RoboDK station: Celda_Soldadura_Estator_Grupo4_v03.rdk

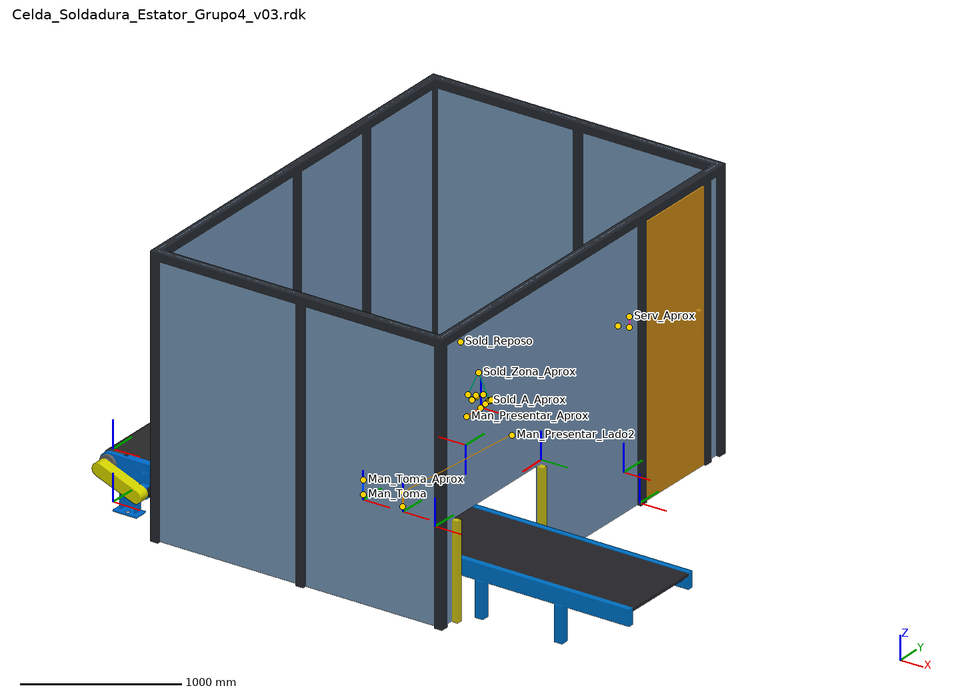
[picture v0: the station drawn from its stored meshes, robots at their saved joint values, targets as dots, program paths as lines]
Station Celda_Soldadura_Estator_Grupo4_v03 (saved by RoboDK 6.1.1). Poses are relative to the parent item; angles as X-Y-Z fixed-axis rotations.
Station parameters (name, value as stored): PIEZA_EN_TOMA, 0, PIEZA_PRESENTADA, 0, ARCO_TIG, 0, SOLDADURA_TERMINADA, 0
  - frame Frame_Celda at (0, 0, 0) mm
    - frame Base_Manipulador_IRB1200 at (0, 0, 0) mm
      - robot ABB IRB 1200-7/0.7: 6 axes, payload 7 kg, reach 703 mm, repeatability 0.02 mm, weight 54 kg
          modified DH rows (alpha deg, a mm, theta deg, d mm): 0, 0, 0, 399; -90, 0, -90, 0; 0, 350, 0, 0; -90, 42, 0, 351; 90, 0, 0, 0; -90, 0, 180, 82
          joint limits [-170, -100, -200, -270, -130, -360] to [170, 135, 70, 270, 130, 360]; home [0, 0, 0, 0, 0, 0]; saved at [0, -20, 30, 0, 80, 0]
        - frame RobotiQ 2F-85 Gripper (Mechanism) Base at (0, 0, 0) mm
          - robot Pinza_2F85 (model RobotiQ 2F85): 1 axes, payload 5 kg
              joint limits [0] to [85]; home [85]; saved at [0]
        - tool TCP_Pinza, TCP at (0, 0, 150) mm
    - frame Base_Soldador_CRB1300 at (0, 1150, 0) mm, rotated rx 0 ry 0 rz -90 deg
      - robot ABB CRB 1300-10/1.15: 6 axes
          modified DH rows (alpha deg, a mm, theta deg, d mm): 0, 0, 0, 544; -90, 150, -90, 0; 0, 575, 0, 0; -90, 40, 0, 425; 90, 0, 0, 0; -90, 0, 180, 90
          joint limits [-180, -95, -210, -230, -130, -242] to [180, 155, 65, 230, 130, 242]; home [0, 0, 0, 0, 0, 0]; saved at [0, -10, 10, 0, 60, 0]
        - tool Antorcha_TIG, TCP at (0, 0, 207) mm, size 80 x 80 x 207 mm, geometry from antorcha_tig.stl
    - frame Base_Cinta_Pasante at (-1830, -860, 0) mm
      - robot Cinta_Pasante: 1 axes
          modified DH rows (alpha deg, a mm, theta deg, d mm): 0, 0, 0, 0 linear
          base shift (0, 0, 0) mm, rotated rx 0 ry 90 rz 0 deg
          joint limits [-900000] to [900000]; home [0]; saved at [0]
        - frame Frame_Banda at (0, 0, 0) mm
          - frame Frame_Piezas_Soldadas at (0, 0, 0) mm
          - object Estator_1 at (1680, 300, 0) mm, size 105 x 105 x 55 mm, geometry from paquete_estator.stl
          - object Estator_2 at (1380, 300, 0) mm, size 105 x 105 x 55 mm, geometry from paquete_estator.stl
          - object Estator_3 at (1080, 300, 0) mm, size 105 x 105 x 55 mm, geometry from paquete_estator.stl
          - object Estator_4 at (780, 300, 0) mm, size 105 x 105 x 55 mm, geometry from paquete_estator.stl
    - object Sensor_Pieza_En_Toma at (-150, -900, 396.5) mm, rotated rx 0 ry 0 rz 90 deg, size 683.3 x 45.2 x 12.5 mm, geometry from Laser-Sensor.stl
    - object Estacion_Servicio_Antorcha at (520, 1300, 0) mm, size 250 x 250 x 1000 mm, geometry from estacion_servicio_antorcha.stl
    - frame Frame_Cerramiento at (0, 0, 0) mm
      - frame Bisagra_Puerta at (850, 1000, 0) mm
        - object Puerta at (0, 0, 0) mm, size 60 x 700 x 1920 mm, geometry from puerta.stl
      - object Cerramiento_Estructura at (0, 0, 0) mm, size 2210 x 3060 x 2000 mm, geometry from cerramiento_estructura_v03.stl
      - object Cerramiento_Paneles at (0, 0, 0) mm, size 2154 x 3004 x 2000 mm, geometry from cerramiento_paneles_v03.stl
      - object Cortina_Luz_Entrada at (-1330, 0, 0) mm, size 40 x 960 x 700 mm, geometry from cortina_luz_cinta.stl
      - object Cortina_Luz_Salida at (880, 0, 0) mm, size 40 x 960 x 700 mm, geometry from cortina_luz_cinta.stl
    - frame Frame_Soldadura at (0, 500, 620) mm
      - target Man_Presentar_Aprox (Cartesian target) at (0, -157.5, 0) mm, rotated rx -90 ry 0 rz 0 deg; joints [0, 0, 0, 0, 0, 0] of ABB IRB 1200-7/0.7
      - target Man_Presentar_Lado1 (Cartesian target) at (0, -7.5, 0) mm, rotated rx -90 ry 0 rz 0 deg; joints [0, 0, 0, 0, 0, 0] of ABB IRB 1200-7/0.7
      - target Man_Presentar_Lado2 (joint target) at (583, -500, 171) mm, rotated rx 0 ry 90 rz 0 deg; joints [90, -11.774, 38.724, 0, -26.95, 90] of ABB IRB 1200-7/0.7
      - target Man_Presentar_Aprox_Lado2 (joint target) at (583, -500, 171) mm, rotated rx 0 ry 90 rz 0 deg; joints [90, -43.636, 55.703, 0, -12.068, 90] of ABB IRB 1200-7/0.7
      - target Sold_Zona_Aprox (Cartesian target) at (0, -26.5, 250) mm, rotated rx 180 ry 0 rz 90 deg; joints [103.36, 41.617, 53.414, 0, -5.031, 103.36] of ABB CRB 1300-10/1.15
      - target Sold_A_Aprox (Cartesian target) at (78.2, -26.5, 78.2) mm, rotated rx -135 ry 0 rz 90 deg; joints [98.688, 74.302, 5.58, 7.491, 55.018, 91.856] of ABB CRB 1300-10/1.15
      - target Sold_A_Inicio (Cartesian target) at (49.91, -26.5, 49.91) mm, rotated rx -135 ry 0 rz 90 deg; joints [98.998, 76.411, 8.063, 8.245, 50.464, 91.119] of ABB CRB 1300-10/1.15
      - target Sold_A_Fin (Cartesian target) at (49.91, 26.5, 49.91) mm, rotated rx -135 ry 0 rz 90 deg; joints [102.751, 76.611, 6.557, 11.474, 51.681, 91.918] of ABB CRB 1300-10/1.15
      - target Sold_Transicion_Medio (Cartesian target) at (0, 26.5, 80) mm, rotated rx 180 ry 0 rz 90 deg; joints [108.748, 65.119, 46.933, 0, -22.052, 108.748] of ABB CRB 1300-10/1.15
      - target Sold_B_Inicio (Cartesian target) at (-49.91, 26.5, 49.91) mm, rotated rx 135 ry 0 rz 90 deg; joints [124.163, 102.688, 60.997, 205.222, 111.278, -54.665] of ABB CRB 1300-10/1.15
      - target Sold_B_Fin (Cartesian target) at (-49.91, -26.5, 49.91) mm, rotated rx 135 ry 0 rz 90 deg; joints [115.401, 107.202, 62.682, 200.569, 120.307, -60.716] of ABB CRB 1300-10/1.15
      - target Sold_B_Retiro (Cartesian target) at (-78.2, -26.5, 78.2) mm, rotated rx 135 ry 0 rz 90 deg; joints [-61.951, -75.264, -208.995, 23.114, 57.885, -82.141] of ABB CRB 1300-10/1.15
      - target Sold_A_Salida (Cartesian target) at (56.57, 26.5, 56.57) mm, rotated rx -135 ry 0 rz 90 deg; joints [102.647, 76.107, 6.003, 11.22, 52.72, 92.165] of ABB CRB 1300-10/1.15
      - target Sold_B_Entrada (Cartesian target) at (-56.57, 26.5, 56.57) mm, rotated rx 135 ry 0 rz 90 deg; joints [124.856, 103.181, 62.152, 205.935, 112.476, -53.248] of ABB CRB 1300-10/1.15
    - frame Frame_Toma_Cinta at (-150, -560, 366.5) mm
      - target Man_Toma_Aprox (Cartesian target) at (0, 0, 135) mm, rotated rx 180 ry 0 rz 0 deg; joints [0, 0, 0, 0, 0, 0] of ABB IRB 1200-7/0.7
      - target Man_Toma (Cartesian target) at (0, 0, 35) mm, rotated rx 180 ry 0 rz 0 deg; joints [0, 0, 0, 0, 0, 0] of ABB IRB 1200-7/0.7
    - frame Frame_Servicio at (520, 1300, 0) mm
      - target Serv_Aprox (Cartesian target) at (0, 60, 1050) mm, rotated rx 180 ry 0 rz 0 deg; joints [-125.65, 36.775, -52.607, 69.175, 38.577, -64.055] of ABB CRB 1300-10/1.15
      - target Serv_Verificacion_TCP (Cartesian target) at (0, 60, 973) mm, rotated rx 180 ry 0 rz 0 deg; joints [-125.65, 36.775, -52.607, 69.175, 38.577, -64.055] of ABB CRB 1300-10/1.15
      - target Serv_Cambio_Tungsteno (Cartesian target) at (0, -65, 1035) mm, rotated rx 180 ry 0 rz 0 deg; joints [-125.65, 36.775, -52.607, 69.175, 38.577, -64.055] of ABB CRB 1300-10/1.15
    - target Man_Reposo (joint target) at (583, 0, 791) mm, rotated rx 0 ry 90 rz 0 deg; joints [0, -20, 30, 0, 80, 0] of ABB IRB 1200-7/0.7
    - target Sold_Reposo (joint target) at (0, 278, 1159) mm, rotated rx 0 ry 90 rz -90 deg; joints [0, -10, 10, 0, 60, 0] of ABB CRB 1300-10/1.15
    - target Pinza_Abierta (joint target) at (536.92, 0, 791) mm, rotated rx 0 ry 90 rz 0 deg; joints [85] of Pinza_2F85
    - target Pinza_Cerrada (joint target) at (536.92, 0, 791) mm, rotated rx 0 ry 90 rz 0 deg; joints [0] of Pinza_2F85
    - target Pinza_Sujeta (joint target) at (536.92, 0, 791) mm, rotated rx 0 ry 90 rz 0 deg; joints [35] of Pinza_2F85
    - target Cinta_Posicion_1 (joint target) at (-1830, -860, 366.5) mm; joints [0] of Cinta_Pasante
    - target Cinta_Posicion_2 (joint target) at (-1830, -860, 366.5) mm; joints [300] of Cinta_Pasante
    - target Cinta_Posicion_3 (joint target) at (-1830, -860, 366.5) mm; joints [600] of Cinta_Pasante
    - target Cinta_Posicion_4 (joint target) at (-1830, -860, 366.5) mm; joints [900] of Cinta_Pasante
    - object Cinta_Salida_Banda at (0, 0, 0) mm, size 1880 x 600 x 20 mm, geometry from cinta_extension_banda.stl
    - object Cinta_Salida_Estructura at (0, 0, 0) mm, size 1880 x 700 x 371.5 mm, geometry from cinta_extension_estructura.stl
    - frame Frame_Deposito_Cinta at (150, -560, 366.5) mm
      - target Man_Deposito_Aprox (Cartesian target) at (0, 0, 135) mm, rotated rx 180 ry 0 rz 0 deg; joints [0, -20, 30, 0, 80, 0] of ABB IRB 1200-7/0.7
      - target Man_Deposito (Cartesian target) at (0, 0, 35) mm, rotated rx 180 ry 0 rz 0 deg; joints [0, -20, 30, 0, 80, 0] of ABB IRB 1200-7/0.7
    - target Cinta_Evacuacion (joint target) at (-1830, -860, 366.5) mm; joints [1750] of Cinta_Pasante
  - program Pinza_Abrir (2 instructions, listed below)
  - program Pinza_Cerrar (2 instructions, listed below)
  - program Pinza_Sujetar (2 instructions, listed below)
  - program Cinta_Avanzar_1 (4 instructions, listed below)
  - program Cinta_Avanzar_2 (4 instructions, listed below)
  - program Cinta_Avanzar_3 (4 instructions, listed below)
  - program Cinta_Avanzar_4 (4 instructions, listed below)
  - program Evento_Tomar_Pieza (2 instructions, listed below)
  - program Evento_Soltar_Pieza (2 instructions, listed below)
  - program Man_Ir_Reposo (4 instructions, listed below)
  - program Man_Tomar_Cinta (16 instructions, listed below)
  - program Man_Presentar_Lado1 (8 instructions, listed below)
  - program Man_Presentar_Lado2 (8 instructions, listed below)
  - program Sold_Ir_Reposo (4 instructions, listed below)
  - program Sold_Par_Cordones (34 instructions, listed below)
  - program Sold_Servicio_Antorcha (10 instructions, listed below)
  - program Sold_Cambio_Tungsteno (8 instructions, listed below)
  - program Inicio_Celda (8 instructions, listed below)
  - program Ciclo_Pieza_1 (9 instructions, listed below)
  - program Ciclo_Pieza_2 (9 instructions, listed below)
  - program Ciclo_Pieza_3 (9 instructions, listed below)
  - program Ciclo_Pieza_4 (9 instructions, listed below)
  - program Fin_Lote (6 instructions, listed below)
  - program Programa_Principal (8 instructions, listed below)
  - program Man_Depositar_Cinta (19 instructions, listed below)
  - program Cinta_Evacuar (2 instructions, listed below)
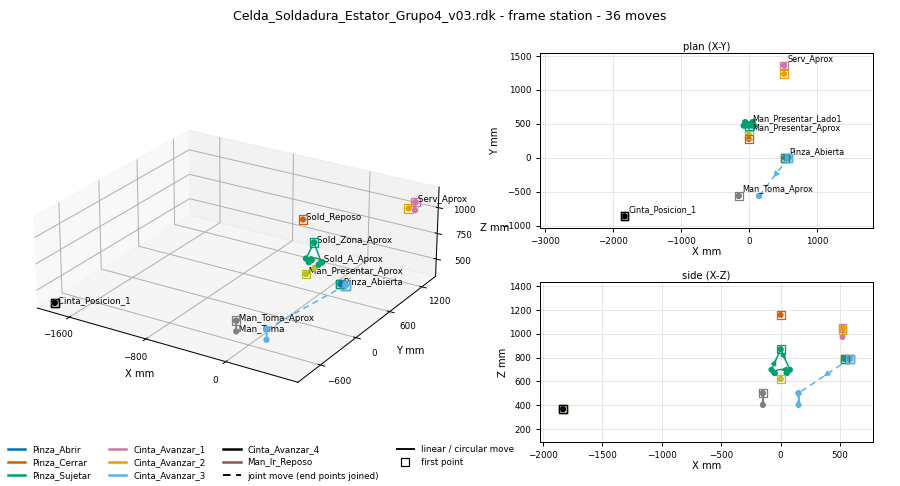
[picture p0: tool path of Celda_Soldadura_Estator_Grupo4_v03.rdk in frame station, 36 of 36 moves have a stored position in this frame; points joined in program order, loops and branches not executed]

--- program Pinza_Abrir (robot Pinza_2F85) ---
  Apertura máxima: reposo de la pinza
  MoveJ (Pinza_Abierta)

--- program Pinza_Cerrar (robot Pinza_2F85) ---
  Dedos juntos para entrar o salir del agujero del estator
  MoveJ (Pinza_Cerrada)

--- program Pinza_Sujetar (robot Pinza_2F85) ---
  Agarre interior: los dedos se abren contra el agujero de Ø55
  MoveJ (Pinza_Sujeta)

--- program Cinta_Avanzar_1 (robot Cinta_Pasante) ---
  Lleva el estator 1 del lote a la posición de toma
  MoveJ (Cinta_Posicion_1)
  Señal del sensor láser: hay pieza en la toma
  Set PIEZA_EN_TOMA=1

--- program Cinta_Avanzar_2 (robot Cinta_Pasante) ---
  Lleva el estator 2 del lote a la posición de toma
  MoveJ (Cinta_Posicion_2)
  Señal del sensor láser: hay pieza en la toma
  Set PIEZA_EN_TOMA=1

--- program Cinta_Avanzar_3 (robot Cinta_Pasante) ---
  Lleva el estator 3 del lote a la posición de toma
  MoveJ (Cinta_Posicion_3)
  Señal del sensor láser: hay pieza en la toma
  Set PIEZA_EN_TOMA=1

--- program Cinta_Avanzar_4 (robot Cinta_Pasante) ---
  Lleva el estator 4 del lote a la posición de toma
  MoveJ (Cinta_Posicion_4)
  Señal del sensor láser: hay pieza en la toma
  Set PIEZA_EN_TOMA=1

--- program Evento_Tomar_Pieza (robot ABB IRB 1200-7/0.7) ---
  Engancha a TCP_Pinza el estator que la pinza acaba de sujetar
  Adjuntar a TCP_Pinza

--- program Evento_Soltar_Pieza (robot ABB IRB 1200-7/0.7) ---
  Libera el estator sobre la banda (Frame_Piezas_Soldadas)
  Separar de TCP_Pinza

--- program Man_Ir_Reposo (robot ABB IRB 1200-7/0.7) ---
  Posición de reposo fuera de la zona de soldadura
  Est. herr: TCP_Pinza
  Establecer velocidad (500.0 mm/s)
  MoveJ (Man_Reposo)

--- program Man_Tomar_Cinta (robot ABB IRB 1200-7/0.7) ---
  Toma el estator de la cinta con agarre interior
  Est. Ref.: Frame_Toma_Cinta
  Est. herr: TCP_Pinza
  Wait PIEZA_EN_TOMA=1
  Establecer velocidad (500.0 mm/s)
  Suave(5)
  MoveJ (Man_Toma_Aprox)
  Llamar Pinza_Cerrar
  Suave(0)
  Establecer velocidad (100.0 mm/s)
  Entrada vertical en el agujero: MoveL para no rozar la pieza
  MoveL (Man_Toma)
  Llamar Pinza_Sujetar
  Llamar Evento_Tomar_Pieza
  Set PIEZA_EN_TOMA=0
  MoveL (Man_Toma_Aprox)

--- program Man_Presentar_Lado1 (robot ABB IRB 1200-7/0.7) ---
  Presenta las aristas A y B arriba, con el eje del estator hacia el soldador
  Est. Ref.: Frame_Soldadura
  Est. herr: TCP_Pinza
  Establecer velocidad (500.0 mm/s)
  MoveJ (Man_Presentar_Aprox)
  Establecer velocidad (100.0 mm/s)
  MoveL (Man_Presentar_Lado1)
  Set PIEZA_PRESENTADA=1

--- program Man_Presentar_Lado2 (robot ABB IRB 1200-7/0.7) ---
  Gira 180° sobre el eje de la pinza (J6) para subir las aristas C y D
  Est. Ref.: Frame_Soldadura
  Est. herr: TCP_Pinza
  Wait SOLDADURA_TERMINADA=1
  Set SOLDADURA_TERMINADA=0
  Establecer velocidad (100.0 mm/s)
  MoveJ (Man_Presentar_Lado2)
  Set PIEZA_PRESENTADA=1

--- program Sold_Ir_Reposo (robot ABB CRB 1300-10/1.15) ---
  Reposo del soldador fuera del volumen de giro de la pieza
  Est. herr: Antorcha_TIG
  Establecer velocidad (500.0 mm/s)
  MoveJ (Sold_Reposo)

--- program Sold_Par_Cordones (robot ABB CRB 1300-10/1.15) ---
  Suelda las dos aristas superiores del estator presentado
  Est. Ref.: Frame_Soldadura
  Est. herr: Antorcha_TIG
  Wait PIEZA_PRESENTADA=1
  Establecer velocidad (500.0 mm/s)
  Suave(5)
  MoveJ (Sold_Zona_Aprox)
  Suave(0)
  Establecer velocidad (100.0 mm/s)
  Aproximación radial a la arista A
  MoveL (Sold_A_Aprox)
  MoveL (Sold_A_Inicio)
  Cordón A: arco encendido, avance recto a velocidad de soldadura
  Set ARCO_TIG=1
  Establecer velocidad (8.0 mm/s)
  MoveL (Sold_A_Fin)
  Set ARCO_TIG=0
  Establecer velocidad (100.0 mm/s)
  Separación radial: la punta sale del escalón antes de rodear la pieza
  MoveL (Sold_A_Salida)
  Transición en arco alrededor del eje del estator, a radio constante
  MoveC (Sold_Transicion_Medio, Sold_B_Entrada)
  MoveL (Sold_B_Inicio)
  Cordón B: avance recto en sentido contrario al A
  Set ARCO_TIG=1
  Establecer velocidad (8.0 mm/s)
  MoveL (Sold_B_Fin)
  Set ARCO_TIG=0
  Establecer velocidad (100.0 mm/s)
  MoveL (Sold_B_Retiro)
  MoveL (Sold_Zona_Aprox)
  Set PIEZA_PRESENTADA=0
  Set SOLDADURA_TERMINADA=1
  Llamar Sold_Ir_Reposo

--- program Sold_Servicio_Antorcha (robot ABB CRB 1300-10/1.15) ---
  Verificación del TCP al final de cada lote
  Est. Ref.: Frame_Servicio
  Est. herr: Antorcha_TIG
  Establecer velocidad (500.0 mm/s)
  MoveJ (Serv_Aprox)
  Establecer velocidad (100.0 mm/s)
  Bajada vertical hasta el cruce de los haces
  MoveL (Serv_Verificacion_TCP)
  MoveL (Serv_Aprox)
  Llamar Sold_Ir_Reposo

--- program Sold_Cambio_Tungsteno (robot ABB CRB 1300-10/1.15) ---
  Cambio o reafilado del tungsteno. Se ejecuta a pedido, con la celda detenida
  Est. Ref.: Frame_Servicio
  Est. herr: Antorcha_TIG
  Establecer velocidad (500.0 mm/s)
  MoveJ (Serv_Cambio_Tungsteno)
  Pausa para el operario: abrir puerta, cambiar electrodo, ajustar saliente
  Parar
  Llamar Sold_Servicio_Antorcha

--- program Inicio_Celda (robot ABB IRB 1200-7/0.7) ---
  Estado inicial conocido: robots en reposo, pinza abierta, arco apagado
  Set ARCO_TIG=0
  Set PIEZA_EN_TOMA=0
  Set PIEZA_PRESENTADA=0
  Set SOLDADURA_TERMINADA=0
  Llamar Sold_Ir_Reposo
  Llamar Man_Ir_Reposo
  Llamar Pinza_Abrir

--- program Ciclo_Pieza_1 (robot ABB IRB 1200-7/0.7) ---
  Ciclo completo del estator 1: tomar, soldar 4 cordones, devolver a la banda
  Llamar Cinta_Avanzar_1
  Llamar Man_Tomar_Cinta
  Llamar Man_Presentar_Lado1
  Llamar Sold_Par_Cordones
  Llamar Man_Presentar_Lado2
  Llamar Sold_Par_Cordones
  Llamar Man_Depositar_Cinta
  Llamar Man_Ir_Reposo

--- program Ciclo_Pieza_2 (robot ABB IRB 1200-7/0.7) ---
  Ciclo completo del estator 2: tomar, soldar 4 cordones, devolver a la banda
  Llamar Cinta_Avanzar_2
  Llamar Man_Tomar_Cinta
  Llamar Man_Presentar_Lado1
  Llamar Sold_Par_Cordones
  Llamar Man_Presentar_Lado2
  Llamar Sold_Par_Cordones
  Llamar Man_Depositar_Cinta
  Llamar Man_Ir_Reposo

--- program Ciclo_Pieza_3 (robot ABB IRB 1200-7/0.7) ---
  Ciclo completo del estator 3: tomar, soldar 4 cordones, devolver a la banda
  Llamar Cinta_Avanzar_3
  Llamar Man_Tomar_Cinta
  Llamar Man_Presentar_Lado1
  Llamar Sold_Par_Cordones
  Llamar Man_Presentar_Lado2
  Llamar Sold_Par_Cordones
  Llamar Man_Depositar_Cinta
  Llamar Man_Ir_Reposo

--- program Ciclo_Pieza_4 (robot ABB IRB 1200-7/0.7) ---
  Ciclo completo del estator 4: tomar, soldar 4 cordones, devolver a la banda
  Llamar Cinta_Avanzar_4
  Llamar Man_Tomar_Cinta
  Llamar Man_Presentar_Lado1
  Llamar Sold_Par_Cordones
  Llamar Man_Presentar_Lado2
  Llamar Sold_Par_Cordones
  Llamar Man_Depositar_Cinta
  Llamar Man_Ir_Reposo

--- program Fin_Lote (robot ABB IRB 1200-7/0.7) ---
  Lote completo: verificación del TCP y evacuación de las piezas soldadas
  Llamar Sold_Servicio_Antorcha
  Llamar Cinta_Evacuar
  Reposición del lote (simula al operario que carga la entrada y retira la salida, afuera)
  Inicio Cinta_Pasante
  Mover objetos

--- program Programa_Principal (robot ABB IRB 1200-7/0.7) ---
  Celda de soldadura TIG de paquetes de estator - Grupo 4
  Un lote = 4 estatores = un pallet. El programa se repite en bucle
  Llamar Inicio_Celda
  Llamar Ciclo_Pieza_1
  Llamar Ciclo_Pieza_2
  Llamar Ciclo_Pieza_3
  Llamar Ciclo_Pieza_4
  Llamar Fin_Lote

--- program Man_Depositar_Cinta (robot ABB IRB 1200-7/0.7) ---
  Devuelve el estator soldado a la banda, aguas abajo de la toma
  Est. Ref.: Frame_Deposito_Cinta
  Est. herr: TCP_Pinza
  Wait SOLDADURA_TERMINADA=1
  Set SOLDADURA_TERMINADA=0
  Establecer velocidad (100.0 mm/s)
  MoveJ (Man_Presentar_Lado2)
  MoveL (Man_Presentar_Aprox_Lado2)
  Establecer velocidad (500.0 mm/s)
  Suave(5)
  MoveJ (Man_Reposo)
  MoveJ (Man_Deposito_Aprox)
  Suave(0)
  Establecer velocidad (100.0 mm/s)
  Bajada vertical hasta apoyar la pieza en la banda
  MoveL (Man_Deposito)
  Llamar Pinza_Cerrar
  Llamar Evento_Soltar_Pieza
  MoveL (Man_Deposito_Aprox)

--- program Cinta_Evacuar (robot Cinta_Pasante) ---
  Avance final: saca el lote soldado por la salida de la celda
  MoveJ (Cinta_Evacuacion)
